CASE eHomeIndexState OF
    E_HomeIndexState.Idle:
        // Wait for homing procedure to be initiated by the drive
        IF rtHomingStart.Q THEN
            Reset();
            bCentered := FALSE;
            // Preserve current velocity for restore after homing, fall back to default
            IF iMotionStage.MotionCmd.fVelocity <> 0.0 THEN
                fPrevVelocity := iMotionStage.MotionCmd.fVelocity;
            ELSE
                fPrevVelocity := fDefaultVelocity;
            END_IF
            eHomeIndexState := E_HomeIndexState.Homing;
        END_IF

    E_HomeIndexState.Homing:
        // Wait for the first rising edge of the index pulse.
        // Transition immediately on detection - HomingUnlatch owns the latch timer,
        // preventing re-entry here and thus ignoring any spurious subsequent pulses.
        IF rtHomePulse.Q THEN
            bHomePulseLatched := TRUE;
            nLatchStartTick := nCurTick;
            iMotionStage.HomeLimit := TRUE;
            eHomeIndexState := E_HomeIndexState.HomingUnlatch;
        END_IF

    E_HomeIndexState.HomingUnlatch:
        // Hold HomeLimit high for nLatchDurationNs to ensure the drive sees the pulse.
        // Any further index pulses are ignored by virtue of being in this state.
        IF (nCurTick - nLatchStartTick) >= nLatchDurationNs THEN
            bHomePulseLatched := FALSE;
            iMotionStage.HomeLimit := FALSE;
            eHomeIndexState := E_HomeIndexState.WaitHomeDone;
        END_IF

    E_HomeIndexState.WaitHomeDone:
        // Index pulse sequence complete. Wait for drive to assert both bDone and
        // bHomed, confirming the homing move has fully settled.
        IF rtWaitHomeIndexDone.Q THEN
            iMotionStage.AbsoluteMoveDefault(
                Position := fCenterOffset,
                Velocity := 15.0,
            );
           eHomeIndexState := E_HomeIndexState.CenterMove;
        END_IF

    E_HomeIndexState.CenterMove:
        // AbsoluteMoveDefault clears bDone before starting, so rtDoneAlign will
        // only fire on the fresh rising edge from this move completing.
        IF rtCenterDone.Q THEN
            // Issue MC_SetPosition to define current position as zero.
            fbMcSetPosition.Execute := TRUE;
            eHomeIndexState := E_HomeIndexState.WaitCenterDone;
        END_IF

    E_HomeIndexState.WaitCenterDone:

        // fbMcSetPosition runs unconditionally below the CASE each cycle.
        IF fbMcSetPosition.Done THEN
            fbMcSetPosition.Execute := FALSE;
            // Position zeroed - mark sequence outputs and advance to Finished
            bCentered := TRUE;
            bHomeDone := TRUE;
            eHomeIndexState := E_HomeIndexState.HomingDone;
        END_IF

    E_HomeIndexState.HomingDone:
        // Restore motion parameters to pre-homing state and enable backlash
        // compensation, then return to Idle ready for next homing cycle.
        bHomePulseLatched := FALSE;
        iMotionStage.SetDefaultMotionParameters(
            HomePosition := 0.0,
            Velocity     := fPrevVelocity,
        );
        eHomeIndexState := E_HomeIndexState.Idle;

    E_HomeIndexState.Error:
        // Latch error output and safe all drive signals.
        // Caller must invoke Reset() to clear and return to Idle.
        bLocalError := TRUE;
        iMotionStage.HomeLimit := FALSE;
        fbMcSetPosition.Execute := FALSE;
        bCentered := FALSE;
        bHomeDone := FALSE;

END_CASE

// MC_SetPosition runs every cycle - Execute is gated by WaitAlignDone state above
fbMcSetPosition(
    Axis     := GVL_AXES.Axes[1],
    Mode     := 0,
    Position := 0.0
);

//FB_Init is always available implicitly and it is used primarily for initialization.
//The return value is not evaluated. For a specific influence, you can also declare the
//methods explicitly and provide additional code there with the standard initialization
//code. You can evaluate the return value.
METHOD FB_Init: BOOL
VAR_INPUT
    bInitRetains: BOOL; // TRUE: the retain variables are initialized (reset warm / reset cold)
    bInCopyCode: BOOL;  // TRUE: the instance will be copied to the copy code afterward (online change)
    iMotionStage : I_MotionStage;
END_VAR
THIS^.iMotionStage := iMotionStage ;
END_METHOD

METHOD Reset
VAR_INPUT
END_VAR
bHomePulseLatched := FALSE;
iMotionStage.HomeLimit := FALSE;
bCentered := FALSE;
bHomeDone := FALSE;
bLocalError := FALSE;
eHomeIndexState := E_HomeIndexState.Idle;
END_METHOD

END_FUNCTION_BLOCK

// ---- POUs/FB_SpindleTaskMonitoring.TcPOU
FUNCTION_BLOCK FB_SpindleTaskMonitoring
VAR_INPUT
    iMotionStage : I_MotionStage; // Interface, assigned via FB_Init at instantiation
END_VAR
VAR_OUTPUT
    nTaskExceedCounter : UDINT;   // Current overrun counter
    nExceedsDelta      : UDINT;   // Difference since last check
    bNewExceeds        : BOOL;    // TRUE if new overrun detected
    bError             : BOOL;    // FB error flag
    nErrorId           : UDINT;   // FB error code
END_VAR
VAR
    fbReadTaskExceedCounter : FB_ReadTaskExceedCounter;
    fBusyEdge               : F_TRIG;
    nPreviousCounter        : UDINT := 0;
    nCurTick                : ULINT := 0;
    nLastCheckTick          : ULINT := 0;
    nCheckIntervalNs        : ULINT := 1_000_000_000; // 1s
    bMonitorRequest         : BOOL := FALSE;
    bFBResetSent            : BOOL := FALSE;
END_VAR

IF (iMotionStage = 0) THEN
    // Outputs default values for fault/no interface assignment
    nTaskExceedCounter := 0;
    nExceedsDelta := 0;
    bNewExceeds := FALSE;
    bError := FALSE;
    nErrorId := 0;
    RETURN;
END_IF

nCurTick := F_GetCurDcTickTime64();

IF (nCurTick - nLastCheckTick) >= nCheckIntervalNs THEN
    bMonitorRequest := TRUE;
    nLastCheckTick := nCurTick;
END_IF

fbReadTaskExceedCounter(
    bExecute := bMonitorRequest,
    nTaskAdsPort := TwinCAT_SystemInfoVarList._TaskInfo[GETCURTASKINDEXEX()].AdsPort
);

fBusyEdge(CLK := fbReadTaskExceedCounter.bBusy);

bError   := fbReadTaskExceedCounter.bError;
nErrorId := fbReadTaskExceedCounter.nErrorId;

IF fBusyEdge.Q AND NOT bError THEN
    nTaskExceedCounter := fbReadTaskExceedCounter.nExceedCounter;
    nExceedsDelta := 0;
    bNewExceeds := FALSE;
    IF nTaskExceedCounter > nPreviousCounter THEN
        bNewExceeds := TRUE;
        nExceedsDelta := nTaskExceedCounter - nPreviousCounter;
        nPreviousCounter := nTaskExceedCounter;

        // Issue spindle reset via the interface
        IF NOT bFBResetSent THEN
            iMotionStage.MotionCmd.bReset := TRUE;
            bFBResetSent := TRUE;
        END_IF
    ELSE
        iMotionStage.MotionCmd.bReset := FALSE;
        bFBResetSent := FALSE;
    END_IF

    bMonitorRequest := FALSE;
END_IF

IF bError THEN
    bMonitorRequest := FALSE;
    nExceedsDelta := 0;
    bNewExceeds := FALSE;
    iMotionStage.MotionCmd.bReset := FALSE;
    bFBResetSent := FALSE;
END_IF

END_FUNCTION_BLOCK
